// TIA Portal project "template" (V17)
// Primeiro projeto de automação industrial utilizando o software TIA17

(* hardware
DEVICE "S7-1500/ET200MP station_1"  S7-1500 station
   slot 0: "Rail_0"  Rack  6ES7 590-1***0-0AA0
   slot 1: "PLC_1"  CPU 1516-3 PN/DP  6ES7 516-3AN01-0AB0  V2.9
      slot 3: "CPU display_1"  6ES7591-1BA00-0AA0
      slot 32768: "PROFINET interface_1"  X1
         slot 32769: "Port_1"  X1 P1
         slot 32770: "Port_2"  X1 P2
      slot 33024: "PROFINET interface_2"  X2
         slot 33025: "Port_1"  X2 P1
      slot 33280: "DP interface_1"  X3
      slot 34817: "Virtual CP interface port_1"  Virtual CP interface port  Virtual CP interface port
   slot 2: "DI 32x24VDC HF_1"  DI 32x24VDC HF  6ES7 521-1BL00-0AB0  V2.1
   slot 3: "DQ 32x24VDC/0.5A HF_1"  DQ 32x24VDC/0.5A HF  6ES7 522-1BL01-0AB0  V1.0
*)

// ===== PLC "PLC_1"  CPU 1516-3 PN/DP =====

VAR_GLOBAL   // PLC tag table "Default tag table"
   "System_Byte" AT %MB1 : Byte;
   "FirstScan" AT %M1.0 : Bool;
   "DiagStatusUpdate" AT %M1.1 : Bool;
   "AlwaysTRUE" AT %M1.2 : Bool;
   "AlwaysFALSE" AT %M1.3 : Bool;
   "Clock_Byte" AT %MB100 : Byte;
   "Clock_10Hz" AT %M100.0 : Bool;
   "Clock_5Hz" AT %M100.1 : Bool;
   "Clock_2.5Hz" AT %M100.2 : Bool;
   "Clock_2Hz" AT %M100.3 : Bool;
   "Clock_1.25Hz" AT %M100.4 : Bool;
   "Clock_1Hz" AT %M100.5 : Bool;
   "Clock_0.625Hz" AT %M100.6 : Bool;
   "Clock_0.5Hz" AT %M100.7 : Bool;
END_VAR

DATA_BLOCK "MDB_RD_CLIENT"   // DB2
{ S7_Optimized_Access := 'TRUE' }
VERSION : 0.1
   VAR
      dadosLeitura : Array[0..70] of Word;
      conexao : TCON_IP_v4;
   END_VAR
BEGIN
   conexao.InterfaceId := 64;
   conexao.ActiveEstablished := true;
   conexao.ID := 1;
   conexao.ConnectionType := 11;
   conexao.RemoteAddress.ADDR[1] := 169;
   conexao.RemoteAddress.ADDR[2] := 254;
   conexao.RemoteAddress.ADDR[3] := 171;
   conexao.RemoteAddress.ADDR[4] := 200;
   conexao.RemotePort := 502;
END_DATA_BLOCK

DATA_BLOCK "MDB_WRITE_ATUADORES"   // DB3
{ S7_Optimized_Access := 'TRUE' }
VERSION : 0.1
   VAR
      dadosEscrita : Array[0..2] of Word;
      conexao : TCON_IP_v4;
   END_VAR
BEGIN
   conexao.InterfaceId := 64;
   conexao.ID := 2;
   conexao.ConnectionType := 11;
   conexao.ActiveEstablished := true;
   conexao.RemoteAddress.ADDR[1] := 169;
   conexao.RemoteAddress.ADDR[2] := 254;
   conexao.RemoteAddress.ADDR[3] := 171;
   conexao.RemoteAddress.ADDR[4] := 200;
   conexao.RemotePort := 502;
END_DATA_BLOCK

DATA_BLOCK "MDB_WRITE_ESTEIRA"   // DB4
{ S7_Optimized_Access := 'TRUE' }
VERSION : 0.1
   VAR
      dadosEscrita : Array[0..1] of Word;
      conexao : TCON_IP_v4;
   END_VAR
BEGIN
   conexao.InterfaceId := 64;
   conexao.ID := 3;
   conexao.ConnectionType := 11;
   conexao.ActiveEstablished := true;
   conexao.RemoteAddress.ADDR[1] := 169;
   conexao.RemoteAddress.ADDR[2] := 254;
   conexao.RemoteAddress.ADDR[3] := 171;
   conexao.RemoteAddress.ADDR[4] := 200;
   conexao.RemotePort := 502;
END_DATA_BLOCK

DATA_BLOCK "MDB_WRITE_SEPARADORES"   // DB5
{ S7_Optimized_Access := 'TRUE' }
VERSION : 0.1
   VAR
      dadosEscrita : Array[0..0] of Word;
      conexao : TCON_IP_v4;
   END_VAR
BEGIN
   conexao.InterfaceId := 64;
   conexao.ID := 4;
   conexao.ConnectionType := 11;
   conexao.ActiveEstablished := true;
   conexao.RemoteAddress.ADDR[1] := 169;
   conexao.RemoteAddress.ADDR[2] := 254;
   conexao.RemoteAddress.ADDR[3] := 171;
   conexao.RemoteAddress.ADDR[4] := 200;
   conexao.RemotePort := 502;
END_DATA_BLOCK

DATA_BLOCK "N1_DB"   // DB6
{ S7_Optimized_Access := 'TRUE' }
VERSION : 0.1
// stored: InstanceOfName N1
"N1"
BEGIN
END_DATA_BLOCK

DATA_BLOCK "DB_Producao_N1"   // DB11
{ S7_Optimized_Access := 'TRUE' }
VERSION : 0.1
   VAR
      contPecasVermelhas : Int;
      contPecasVerdes : Int;
      contPecasAmarelas : Int;
      contPecasTotal : Int;
   END_VAR
BEGIN
END_DATA_BLOCK

// folder: System blocks/Program resources

DATA_BLOCK "C1"   // DB1
{ S7_Optimized_Access := 'TRUE' }
AUTHOR : Simatic
FAMILY : IEC
NAME : CNTR
VERSION : 1.0
// stored: InstanceOfName IEC_COUNTER
"IEC_COUNTER"
BEGIN
END_DATA_BLOCK

// folder: (top level)

FUNCTION_BLOCK "N1"   // FB1, SCL
{ S7_Optimized_Access := 'TRUE' }
VERSION : 0.1
   VAR_INPUT
      posAtualX : Int;
      yAv : Bool;
      yRec : Bool;
      zAv : Bool;
      zRec : Bool;
      pcEsteira : Bool;
      pcRampaVerm : Bool;
      pcRampaVerde : Bool;
      pcRampaAmar : Bool;
      corVerm : Bool;
      corVerde : Bool;
      corAmar : Bool;
      SepVermRec : Bool;
      SepVermAv : Bool;
      SepVerdeAv : Bool;
      SepVerdeRec : Bool;
      SepAmarAv : Bool;
      SepAmarRec : Bool;
      chaveGeral : Bool;
      Emerg : Bool;
      start : Bool;
      stop : Bool;
   END_VAR
   VAR_OUTPUT
      velocEst : Int;
      estAvancar : Bool;
      estRecuar : Bool;
      sepVermRecuar : Bool;
      sepVermAvancar : Bool;
      sepVerdeRecuar : Bool;
      sepVerdeAvancar : Bool;
      sepAmarRecuar : Bool;
      sepAmarAvancar : Bool;
      estado : Int;
   END_VAR
   VAR
      tempoDeslocamento : Time;
      qtdTotal : Int;
      qtdAmar : Int;
      qtdVerde : Int;
      corMemorizada : Int;
      qtdVerm : Int;
   END_VAR
BEGIN
   // ==========================================
   // AÇÕES
   // ==========================================
   CASE #estado OF
       0:  // ESTADO INICIAL / RESET / EMERGÊNCIA
           #estAvancar := 0;
           #estRecuar := 0;
           #velocEst := 0;
           #sepVerdeAvancar := 0;
           #sepVerdeRecuar := 1;
           #sepVermAvancar := 0;
           #sepVermRecuar := 1;
           #sepAmarAvancar := 0;
           #sepAmarRecuar := 1;

       1:  // CONDIÇÕES INICIAIS OK (Aguardando Start)
           #sepVerdeRecuar := 0;
           #sepVermRecuar := 0;
           #sepAmarRecuar := 0;
           #velocEst := 0;
           #estAvancar := 0;

       2:  // ESTEIRA RODANDO / PROCURANDO PEÇA (Todos os pistões recuados)
           #velocEst := 60;
           #estAvancar := 1;
           #sepAmarAvancar := 0;
           #sepAmarRecuar := 1;
           #sepVermAvancar := 0;
           #sepVermRecuar := 1;
           #sepVerdeAvancar := 0;
           #sepVerdeRecuar := 1;

       3:  // DESVIADOR AMARELO ABERTO (Aguardando peça entrar na rampa)
           #velocEst := 60;
           #estAvancar := 1;
           #sepAmarRecuar := 0;
           #sepAmarAvancar := 1;

       4:  // DESVIADOR VERMELHO ABERTO (Aguardando peça entrar na rampa)
           #velocEst := 60;
           #estAvancar := 1;
           #sepVermRecuar := 0;
           #sepVermAvancar := 1;

       5:  // DESVIADOR VERDE ABERTO (Aguardando peça entrar na rampa)
           #velocEst := 60;
           #estAvancar := 1;
           #sepVerdeRecuar := 0;
           #sepVerdeAvancar := 1;
   END_CASE;

   // ==========================================
   // TRANSIÇÕES DE ESTADOS
   // ==========================================
   IF #estado = 0 AND #SepAmarRec AND #SepVerdeRec AND #SepVermRec AND #chaveGeral AND NOT #Emerg THEN
       #estado := 1;
   END_IF;

   IF #estado = 1 AND #start AND #chaveGeral AND NOT #Emerg THEN
       #estado := 2;
   END_IF;

   // Detectou a cor -> abre o desviador IMEDIATAMENTE
   IF #estado = 2 AND #corAmar AND #chaveGeral AND NOT #Emerg THEN
       #estado := 3;
   END_IF;

   IF #estado = 2 AND #corVerm AND #chaveGeral AND NOT #Emerg THEN
       #estado := 4;
   END_IF;

   IF #estado = 2 AND #corVerde AND #chaveGeral AND NOT #Emerg THEN
       #estado := 5;
   END_IF;

   // Peça entrou na rampa -> conta e recua o desviador voltando para o estado 2
   IF #estado = 3 AND #pcRampaAmar THEN
       #qtdAmar := #qtdAmar + 1;
       #qtdTotal := #qtdAmar + #qtdVerm + #qtdVerde;
       #estado := 2;
   END_IF;

   IF #estado = 4 AND #pcRampaVerm THEN
       #qtdVerm := #qtdVerm + 1;
       #qtdTotal := #qtdAmar + #qtdVerm + #qtdVerde;
       #estado := 2;
   END_IF;

   IF #estado = 5 AND #pcRampaVerde THEN
       #qtdVerde := #qtdVerde + 1;
       #qtdTotal := #qtdAmar + #qtdVerm + #qtdVerde;
       #estado := 2;
   END_IF;

   "DB_Producao_N1".contPecasVermelhas := #qtdVerm;
   "DB_Producao_N1".contPecasVerdes := #qtdVerde;
   "DB_Producao_N1".contPecasAmarelas := #qtdAmar;
   "DB_Producao_N1".contPecasTotal := #qtdTotal;

   // ==========================================
   // INTERRUPÇÕES DE SEGURANÇA
   // ==========================================
   IF #Emerg OR NOT #chaveGeral OR #stop THEN
       #estado := 0;
   END_IF;
END_FUNCTION_BLOCK

ORGANIZATION_BLOCK "Main"   // OB1, LAD, ProgramCycle
TITLE = "Main Program Sweep (Cycle)"
{ S7_Optimized_Access := 'TRUE' }
VERSION : 0.1
   VAR_INPUT
      Initial_Call : Bool;   // Initial call of this OB
      Remanence : Bool;   // =True, if remanent data are available
   END_VAR
BEGIN

REGION Network 1 (SCL)
   "C1".CTU(CU:="Clock_2Hz", R:="C1".QU, PV:=5);
END_REGION

REGION Network 2
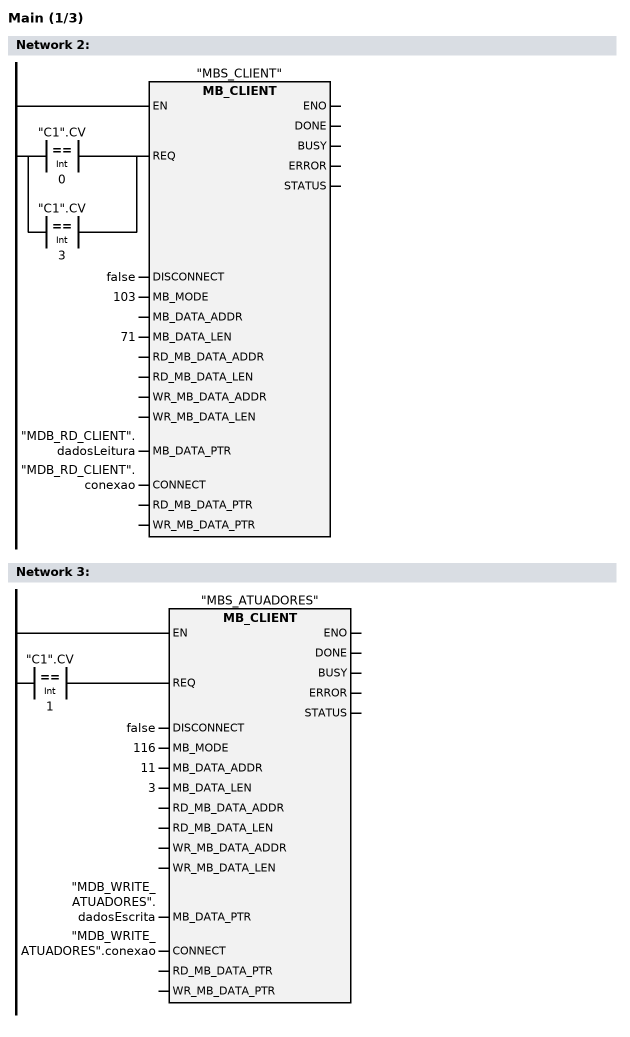
   "MBS_CLIENT"(REQ := ("C1".CV = 0) OR ("C1".CV = 3),   // MB_CLIENT
                DISCONNECT := false,
                MB_MODE := 103,
                MB_DATA_LEN := 71,
                MB_DATA_PTR := "MDB_RD_CLIENT".dadosLeitura,
                CONNECT := "MDB_RD_CLIENT".conexao);
END_REGION

REGION Network 3
   "MBS_ATUADORES"(REQ := "C1".CV = 1,   // MB_CLIENT
                   DISCONNECT := false,
                   MB_MODE := 116,
                   MB_DATA_ADDR := 11,
                   MB_DATA_LEN := 3,
                   MB_DATA_PTR := "MDB_WRITE_ATUADORES".dadosEscrita,
                   CONNECT := "MDB_WRITE_ATUADORES".conexao);
END_REGION

REGION Network 4
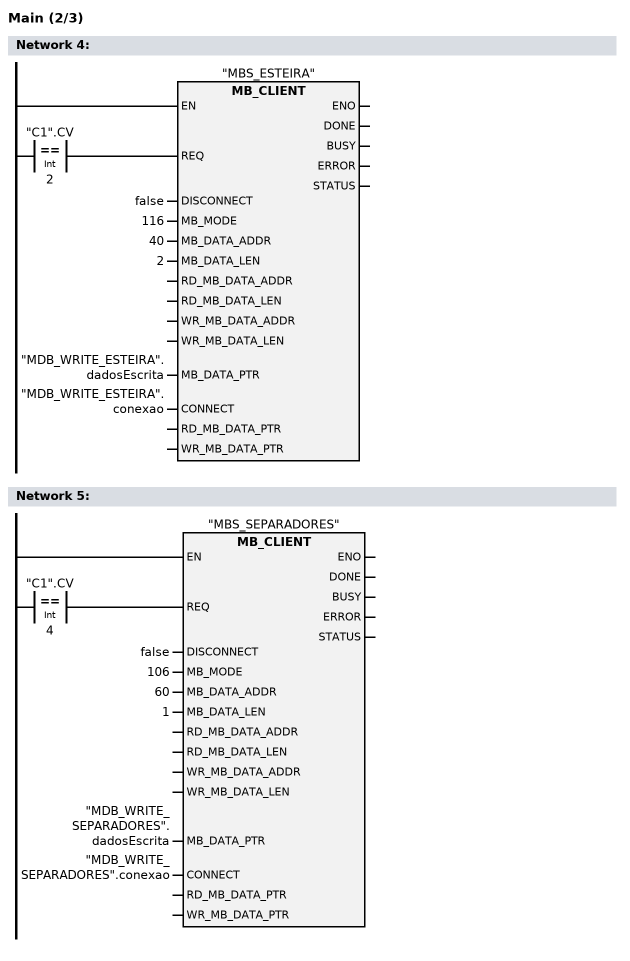
   "MBS_ESTEIRA"(REQ := "C1".CV = 2,   // MB_CLIENT
                 DISCONNECT := false,
                 MB_MODE := 116,
                 MB_DATA_ADDR := 40,
                 MB_DATA_LEN := 2,
                 MB_DATA_PTR := "MDB_WRITE_ESTEIRA".dadosEscrita,
                 CONNECT := "MDB_WRITE_ESTEIRA".conexao);
END_REGION

REGION Network 5
   "MBS_SEPARADORES"(REQ := "C1".CV = 4,   // MB_CLIENT
                     DISCONNECT := false,
                     MB_MODE := 106,
                     MB_DATA_ADDR := 60,
                     MB_DATA_LEN := 1,
                     MB_DATA_PTR := "MDB_WRITE_SEPARADORES".dadosEscrita,
                     CONNECT := "MDB_WRITE_SEPARADORES".conexao);
END_REGION

REGION Network 6
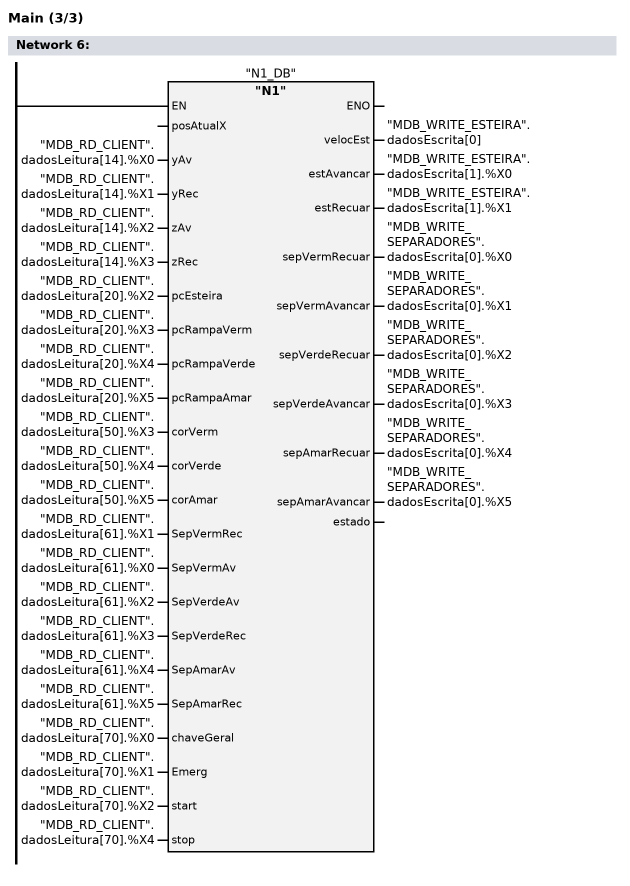
   RUNG wire#powerrail
      "N1_DB"(posAtualX :=, yAv := "MDB_RD_CLIENT".dadosLeitura[14].%X0, yRec := "MDB_RD_CLIENT".dadosLeitura[14].%X1, zAv := "MDB_RD_CLIENT".dadosLeitura[14].%X2, zRec := "MDB_RD_CLIENT".dadosLeitura[14].%X3, pcEsteira := "MDB_RD_CLIENT".dadosLeitura[20].%X2, pcRampaVerm := "MDB_RD_CLIENT".dadosLeitura[20].%X3, pcRampaVerde := "MDB_RD_CLIENT".dadosLeitura[20].%X4, pcRampaAmar := "MDB_RD_CLIENT".dadosLeitura[20].%X5, corVerm := "MDB_RD_CLIENT".dadosLeitura[50].%X3, corVerde := "MDB_RD_CLIENT".dadosLeitura[50].%X4, corAmar := "MDB_RD_CLIENT".dadosLeitura[50].%X5, SepVermRec := "MDB_RD_CLIENT".dadosLeitura[61].%X1, SepVermAv := "MDB_RD_CLIENT".dadosLeitura[61].%X0, SepVerdeAv := "MDB_RD_CLIENT".dadosLeitura[61].%X2, SepVerdeRec := "MDB_RD_CLIENT".dadosLeitura[61].%X3, SepAmarAv := "MDB_RD_CLIENT".dadosLeitura[61].%X4, SepAmarRec := "MDB_RD_CLIENT".dadosLeitura[61].%X5, chaveGeral := "MDB_RD_CLIENT".dadosLeitura[70].%X0, Emerg := "MDB_RD_CLIENT".dadosLeitura[70].%X1, start := "MDB_RD_CLIENT".dadosLeitura[70].%X2, stop := "MDB_RD_CLIENT".dadosLeitura[70].%X4, velocEst => "MDB_WRITE_ESTEIRA".dadosEscrita[0], estAvancar => "MDB_WRITE_ESTEIRA".dadosEscrita[1].%X0, estRecuar => "MDB_WRITE_ESTEIRA".dadosEscrita[1].%X1, sepVermRecuar => "MDB_WRITE_SEPARADORES".dadosEscrita[0].%X0, sepVermAvancar => "MDB_WRITE_SEPARADORES".dadosEscrita[0].%X1, sepVerdeRecuar => "MDB_WRITE_SEPARADORES".dadosEscrita[0].%X2, sepVerdeAvancar => "MDB_WRITE_SEPARADORES".dadosEscrita[0].%X3, sepAmarRecuar => "MDB_WRITE_SEPARADORES".dadosEscrita[0].%X4, sepAmarAvancar => "MDB_WRITE_SEPARADORES".dadosEscrita[0].%X5, estado =>)
   END_RUNG
   // the same network as SCL:
   "N1_DB"(yAv := "MDB_RD_CLIENT".dadosLeitura[14].%X0,   // "N1"
           yRec := "MDB_RD_CLIENT".dadosLeitura[14].%X1,
           zAv := "MDB_RD_CLIENT".dadosLeitura[14].%X2,
           zRec := "MDB_RD_CLIENT".dadosLeitura[14].%X3,
           pcEsteira := "MDB_RD_CLIENT".dadosLeitura[20].%X2,
           pcRampaVerm := "MDB_RD_CLIENT".dadosLeitura[20].%X3,
           pcRampaVerde := "MDB_RD_CLIENT".dadosLeitura[20].%X4,
           pcRampaAmar := "MDB_RD_CLIENT".dadosLeitura[20].%X5,
           corVerm := "MDB_RD_CLIENT".dadosLeitura[50].%X3,
           corVerde := "MDB_RD_CLIENT".dadosLeitura[50].%X4,
           corAmar := "MDB_RD_CLIENT".dadosLeitura[50].%X5,
           SepVermRec := "MDB_RD_CLIENT".dadosLeitura[61].%X1,
           SepVermAv := "MDB_RD_CLIENT".dadosLeitura[61].%X0,
           SepVerdeAv := "MDB_RD_CLIENT".dadosLeitura[61].%X2,
           SepVerdeRec := "MDB_RD_CLIENT".dadosLeitura[61].%X3,
           SepAmarAv := "MDB_RD_CLIENT".dadosLeitura[61].%X4,
           SepAmarRec := "MDB_RD_CLIENT".dadosLeitura[61].%X5,
           chaveGeral := "MDB_RD_CLIENT".dadosLeitura[70].%X0,
           Emerg := "MDB_RD_CLIENT".dadosLeitura[70].%X1,
           start := "MDB_RD_CLIENT".dadosLeitura[70].%X2,
           stop := "MDB_RD_CLIENT".dadosLeitura[70].%X4,
           velocEst => "MDB_WRITE_ESTEIRA".dadosEscrita[0],
           estAvancar => "MDB_WRITE_ESTEIRA".dadosEscrita[1].%X0,
           estRecuar => "MDB_WRITE_ESTEIRA".dadosEscrita[1].%X1,
           sepVermRecuar => "MDB_WRITE_SEPARADORES".dadosEscrita[0].%X0,
           sepVermAvancar => "MDB_WRITE_SEPARADORES".dadosEscrita[0].%X1,
           sepVerdeRecuar => "MDB_WRITE_SEPARADORES".dadosEscrita[0].%X2,
           sepVerdeAvancar => "MDB_WRITE_SEPARADORES".dadosEscrita[0].%X3,
           sepAmarRecuar => "MDB_WRITE_SEPARADORES".dadosEscrita[0].%X4,
           sepAmarAvancar => "MDB_WRITE_SEPARADORES".dadosEscrita[0].%X5);
END_REGION
END_ORGANIZATION_BLOCK